// TIA Portal V20 export
// export: Created 2026-10-20T12:46:28.7864157Z, ExportSetting WithDefaults, DisplayName Totally Integrated Automation Portal, DisplayVersion V20 Update 6, DisplayName TIA Portal Openness, DisplayVersion V20 Update 6, DisplayName TIA Portal Version Control Interface, DisplayVersion V20 Update 6, DisplayName SINAMICS Startdrive Advanced, DisplayVersion V20 SP1, DisplayName SINAMICS Startdrive G130, G150, S120, S150, SINAMICS MV, G220, S200, S210, DisplayVersion V20 SP1, DisplayName SINAMICS Startdrive G110M, G120, G120C, G120D, G120P, G115D, DisplayVersion V20 SP1, DisplayName STEP 7 Professional, DisplayVersion V20 Update 6, DisplayName STEP 7 Safety, DisplayVersion V20 Update 2, DisplayName WinCC Basic/Comfort/Advanced, DisplayVersion V20 Update 6, DisplayName WinCC Unified, DisplayVersion V20 Update 6
DATA_BLOCK "VTD_HMI"   // DB57
{ S7_Optimized_Access := 'TRUE' }
VERSION : 0.1
// stored: AutoNumber true, DBAccessibleFromOPCUA true, IsOnlyStoredInLoadMemory false, IsRetainMemResEnabled false, IsWriteProtectedInAS false, MemoryReserve 100
   VAR
      Start_InBarcodeStation : Array[1..5] of Bool;
      Move_To_Level : Array[1..5] of UInt;
      Mode_Change : Array[1..5] of UInt;
      Manual_Down : Array[1..5] of Bool;
      Pallet_Type : Array[1..5] of UInt;
      Manual_Up : Array[1..5] of Bool;
      Task_ID : Array[1..5] of UInt;
      Reset : Array[1..5] of Bool;
      Enable : Array[1..5] of Bool;
      Progress : Array[1..5] of Int;
      Stop : Array[1..5] of Bool;
      Manual_DP_Extend : Array[1..5] of Bool;
      Manual_DP_Retract : Array[1..5] of Bool;
      ID : Array[1..5] of UInt;
      Cnv_Occupied : Array[1..5] of Bool;
      Motor_Status : Array[1..5] of UInt;
      ID_OLD : Array[1..5] of UInt;
      LE_Error : Array[1..5] of Bool;
      Mode : Array[1..5] of UInt;
      Encoder_Delta : Array[1..5] of Real;
      Warning : Array[1..5] of Bool;
      Current_Level : Array[1..5] of UInt;
      Error : Array[1..5] of Bool;
      Current_Task_ID : Array[1..5] of UInt;
      Pallet_Loaded : Array[1..5] of UInt;
      Stopped : Array[1..5] of Bool;
      SM_State : Array[1..5] of UInt;
      Shuttle_Loaded : Array[1..5] of UInt;
      DP_State : Array[1..5] of UInt;
      AE : Array[1..5] of Real;
      Docked : Array[1..5] of Bool;
      AE_Error : Array[1..5] of Bool;
      Enabled : Array[1..5] of Bool;
      Current_Task_Type : Array[1..5] of UInt;
      Running : Array[1..5] of Bool;
      LE : Array[1..5] of Real;
      Motor_Actual_Speed : Array[1..5] of UInt;
      Motor_SetPoint : Array[1..5] of UInt;
      Motor_Actual_Current : Array[1..5] of Real;
      Motor_Ready : Array[1..5] of Bool;
      "Chain Slack 1" : Array[1..5] of Bool;
      "Chain Slack 3" : Array[1..5] of Bool;
      "Chain Slack 2" : Array[1..5] of Bool;
      "Chain Slack 4" : Array[1..5] of Bool;
      Safety_OK : Array[1..5] of Bool;
      Moving_To_Level : Array[1..5] of UInt;
      Speed_mm_s : Array[1..5] of Real;
      Level_Below_Extractor : Array[1..5] of UInt;
      Actual_Torque : Array[1..5] of UInt;
      DP1_Retracted : Array[1..5] of Bool;
      DP2_Extended : Array[1..5] of Bool;
      Upper_Overtravel : Array[1..5] of Bool;
      DP1_Extended : Array[1..5] of Bool;
      DP2_Retracted : Array[1..5] of Bool;
      Lower_Overtravel : Array[1..5] of Bool;
      Level_Detect1 : Array[1..5] of Bool;
      Lower_Limit : Array[1..5] of Bool;
      Ultimate_Creep : Array[1..5] of Bool;
      Upper_Limet : Array[1..5] of Bool;
      Level_Detect2 : Array[1..5] of Bool;
      Ultimate_Slow : Array[1..5] of Bool;
      Charge_VTD_Commands : Array[1..5] of Bool;
      LE_Bypass : Array[1..5] of Bool;
      Charge_VTD : Array[1..5] of Bool;
   END_VAR
BEGIN
END_DATA_BLOCK
